# EPICS autosave request: soft_iocs/bleps/iocBoot/ioc18id/auto_positions.req
file built_positions.req P=$(P)
